Fanuc KAREL source: kt00726.KL

PROGRAM KT00726
%STACKSIZE=65535
%PRIORITY=65535
%NOLOCKGROUP
VAR
V1 : VECTOR
V2 : VECTOR
OUT : BOOLEAN
BEGIN
V1.X=1.0
V2.Y=2.0
V1.X=1.0
V2.Y=2.0
-- UNRESOLVED_PC line 12 opcodes [22 63 23] marker_code=80
END KT00726
